FUNCTION_BLOCK FB_Temperature
(*

The function block used to control temperature.

Constructor: 		Patryk Panylo
Company:		E. Riexinger GmbH
Date:			23.04.2015
Version:			1.00

Date:			Revision:		Who:				Comment
dd.mm.yyyy		x.xx			Initials			comment

*)
VAR_INPUT
	(* Input variables / Eingang Variablen *)
	bEnable					:BOOL;						(* Enable FB signal *)
	bIn						:BOOL;						(* Input signal *)
	tTimeOut					:TIME := t#5s;					(* Timeout *)
END_VAR
VAR_OUTPUT
	(* Output variables / Ausgang Variablen *)
	bOut					:BOOL;						(* Air pressure ok *)
	bError					:BOOL;						(* Error by no air pressure *)
	bWarning				:BOOL;						(* Warning by no temperature *)
	udnErrorNo				:UDINT;
	udnMessageNo			:UDINT;
	sMsg					:STRING;
END_VAR
VAR_IN_OUT

END_VAR
VAR
	(* Enummerations *)

	(* Variables *)
	bFirstTime				:BOOL;						(* First cycle *)

	(* References *)

	(* Interfaces *)

	(* Instances *)
	tonWatchDog				:TON;						(* Timer to delay *)
END_VAR

IF NOT bEnable
THEN
	bOut := TRUE;
	bError := FALSE;
	udnErrorNo := 0;
	udnMessageNo := 0;
	sMsg := '';
	tonWatchDog(IN := FALSE,
	             		 PT := tTimeOut);
	bFirstTime := FALSE;
	RETURN;
END_IF;

IF NOT bFirstTime
THEN
	bError := FALSE;
	udnErrorNo := 0;
	udnMessageNo := 0;
	sMsg := '';
	tonWatchDog(IN := FALSE,
	             		 PT := tTimeOut);
	bFirstTime := TRUE;
END_IF;

(* Timer starts when came rising edge of signal *)
tonWatchDog(
	IN := NOT bIn,
	PT := tTimeOut
);

bOut := bIn;
bError := NOT bOut
	        AND tonWatchDog.Q;
bWarning := NOT bError
		      AND NOT bOut;

IF NOT bOut
THEN
	IF tonWatchDog.Q                       		 (* Error if air pressure not present *)
	THEN
		udnErrorNo := 1;
		udnMessageNo := 0;
		sMsg := 'Temperature not ok';
	END_IF;
ELSE
	udnErrorNo := 0;
	udnMessageNo := 0;
	sMsg := '';
END_IF;

END_FUNCTION_BLOCK

(* stored: Version 1.1.0.1, ProductVersion 3.1.4024.15
   POU FB_Temperature: Id {f1219414-451d-408a-82ab-eaab5cfbbfd7}, SpecialFunc None *)
